Fanuc KAREL source: kt00748.KL

-- PROVISIONAL review KL for V770-1; original PC SHA256 240073d6d81c35b4b595e4cefcfbdf6d724f3a6e5e08788fa2ec6bc18ec9c4c1
-- Incomplete behavior may be omitted. Consult companion uncertainty JSON. Do not deploy.
PROGRAM KT00748
%NOLOCKGROUP
VAR
  I1 : INTEGER
  I2 : INTEGER
  OUT : INTEGER
BEGIN
  -- UNRESOLVED_PC offsets 5-16; opcodes 2E,23
  -- UNRESOLVED_PC offsets 21-32; opcodes 2E,23
  -- UNRESOLVED_PC offsets 37-48; opcodes 2E,23
  -- UNRESOLVED_PC offsets 53-64; opcodes 2E,23
  -- UNRESOLVED_PC offsets 69-82; opcodes 21,50,23
  -- UNRESOLVED_PC offsets 87-91; opcodes 7F
END KT00748
